FUNCTION_BLOCK FB_EL3356ChannelDiagnosis_1
VAR_INPUT
	stChannelState				:ST_EL3356ChannelState;
END_VAR
VAR_OUTPUT
	bChannelOK					:BOOL;
	bCalibrationInProgress			:BOOL;
END_VAR
VAR

END_VAR


(* General Channel Status *)
IF stChannelState.bOverrange = 0
    AND stChannelState.bError = 0
    AND stChannelState.bSyncError = 0
THEN
	bChannelOK := TRUE;
ELSE
	bChannelOK := FALSE;
END_IF

bCalibrationInProgress := stChannelState.bCalibrationInProgress;

END_FUNCTION_BLOCK

(* stored: Version 1.1.0.1, ProductVersion 3.1.4024.15
   POU FB_EL3356ChannelDiagnosis_1: Id {21217628-b136-4eeb-9174-6ca91da6d694}, SpecialFunc None *)
